TYPE ET_BOSCH_AxisSetLimits :
(
	eWaitExecute := 0,
	eSetReferenceSystem,
	eSetPositionBias,
	eSetLimitPos,
	eWfSetLimitPos,
	eSetLimitNeg,
	eWfSetLimitNeg,
	eEnableLimitPos,
	eWfEnableLimitPos,
	eEnableLimitNeg,
	eWfEnableLimitNeg,
	eEnablePosLagMonitoring,
	eWfEnablePosLagMonitoring,
	eDone := 197,
	eError := 198,
	eNoExecute := 199
);
END_TYPE

(* stored: Version 1.1.0.1, ProductVersion 3.1.4024.15
   DUT ET_BOSCH_AxisSetLimits: Id {db9230c3-db39-45e1-98b0-9fc4d233ea4a} *)
